SUBAPPLICATION SubApp_PC_A (* Geraet A: Objekte/Variablen per PUBLISH_0: I1 CREATE_OBJECT, I2 CREATE_VARIABLE, I3 DELETE_VARIABLE, I4 DELETE_OBJECT *)
  (* Standard: 61499-2; Description: Copyright (c) 2026 Meisterschulen am Ostbahnhof This program and the accompanying materials are made available under the terms of the Eclipse Public License 2.0 which is available at https://www.eclipse.org/legal/epl-2.0/ SPDX-License-Identifier: EPL-2.0 *)
  (* Version 1.0, 2026-10-18, Franz Höpfinger, Meisterschulen am Ostbahnhof, opcua.adoc-Beispiel auf zwei Geraeten *)
  PACKAGE subapp::Training_18_OPC_UA_RES;
  IMPORT VV::const::OPC_UA::myOpcUaAddresses::T18_VAR_CLIENT_READ;
  IMPORT logiBUS::io::DI::logiBUS_DI::Input_I1;
  IMPORT logiBUS::io::DI::logiBUS_DI_Events::BUTTON_PRESS_DOWN;
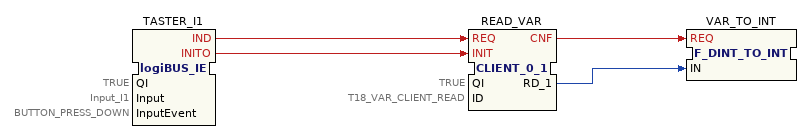
  FBS
    TASTER_I1 : logiBUS::io::DI::logiBUS_IE(QI := TRUE, Input := Input_I1, InputEvent := BUTTON_PRESS_DOWN);
    READ_VAR : iec61499::net::CLIENT_0_1(QI := TRUE, ID := T18_VAR_CLIENT_READ);
    VAR_TO_INT : iec61131::conversion::F_DINT_TO_INT;
  END_FBS
  EVENT_CONNECTIONS
    TASTER_I1.IND TO READ_VAR.REQ;
    TASTER_I1.INITO TO READ_VAR.INIT;
    READ_VAR.CNF TO VAR_TO_INT.REQ;
  END_CONNECTIONS
  DATA_CONNECTIONS
    READ_VAR.RD_1 TO VAR_TO_INT.IN;
  END_CONNECTIONS
END_SUBAPPLICATION
